{attribute 'linkalways'}
{attribute 'no_explicit_call' := 'This FB is a CLASS and must be accessed using methods or properties'}
{attribute 'enable_dynamic_creation'}
FUNCTION_BLOCK Node_F_VN_TransformIntoDisplayableImageExp2 EXTENDS VisionNode
VAR
    ipSrcImage : _ITcVnImage;
    ipDestImage : _ITcVnDisplayableImage;
    bAllowDeepCopy : _BOOL(FALSE);
    nTimestamp : _LINT(0);
    hrPrev : _HRESULT(S_OK);
    hresult : _HRESULT(S_OK);
END_VAR

METHOD PUBLIC Clone : I_Node
VAR
    pNode : POINTER TO Node_F_VN_TransformIntoDisplayableImageExp2;
END_VAR
pNode := __NEW(Node_F_VN_TransformIntoDisplayableImageExp2);
Clone := pNode^;
END_METHOD

METHOD FB_init : BOOL
VAR_INPUT
    bInitRetains : BOOL;
    bInCopyCode : BOOL;
END_VAR
AddInput('ipSrcImage', ipSrcImage);
AddParameter('bAllowDeepCopy', bAllowDeepCopy);
AddParameter('nTimestamp', nTimestamp);
AddInput('hrPrev', hrPrev);
AddOutput('ipDestImage', ipDestImage);
AddOutput('hresult', hresult);
END_METHOD

METHOD PROTECTED OnExecute
hresult.Value := F_VN_TransformIntoDisplayableImageExp2(
    ipSrcImage := ipSrcImage.Value,
    ipDestImage := ipDestImage.Value,
    bAllowDeepCopy := bAllowDeepCopy.Value,
    nTimestamp := nTimestamp.Value,
    hrPrev := hrPrev.Value);
END_METHOD

METHOD PUBLIC PreExecutionCheck
VAR_INPUT
    Check : I_PreExecutionChecks;
END_VAR
Check.IsTrue(ipSrcImage.IsValid, 'ipSrcImage must contain an image');
END_METHOD

END_FUNCTION_BLOCK

(* stored: Version 1.1.0.1, ProductVersion 3.1.4026.19
   POU Node_F_VN_TransformIntoDisplayableImageExp2: Id {36f7be24-4e41-49cd-aa46-ad55d684f65e}, SpecialFunc None
   Folder Constructor: Id {40591ef4-506c-4b9d-ac5f-d3b4b8cfa2b4}
   Method Clone: Id {f906662b-1ecd-404f-a9cd-8fb853f3f4d9}
   Method FB_init: Id {49dcad6f-9956-4cf3-92d3-4f70884f9055}
   Method OnExecute: Id {ccc1d886-8d68-4065-8ca8-d1ac52e0d737}
   Method PreExecutionCheck: Id {0d203290-9227-412e-b5a5-90feee246843} *)
